// TIA Portal V21 export
// export: Created 2026-10-14T03:11:19.0543245Z, ExportSetting WithDefaults, DisplayName Totally Integrated Automation Portal, DisplayVersion V21, DisplayName STEP 7 Professional, DisplayVersion V21, DisplayName STEP 7 Safety, DisplayVersion V21, DisplayName Tech WebApplication, DisplayVersion V21, DisplayName WinCC Basic/Comfort/Advanced, DisplayVersion V21, DisplayName WinCC Unified, DisplayVersion V21
TagTable "PID_LCCA"
  LLCCA_PID_DB_Input : Real  (HMI_Connection_1, 100 ms)
  LLCCA_PID_DB_Out : Real  (HMI_Connection_1, 100 ms)
  LLCCA_PID_DB_Setpoint : Real  (HMI_Connection_1, 100 ms)
  LLCCA_PID_DB_ioKp : Real  (HMI_Connection_1, 1 s)
  LLCCA_PID_DB_ioTi : Real  (HMI_Connection_1, 1 s)
  LLCCA_PID_DB_ioTd : Real  (HMI_Connection_1, 1 s)
  LLCCA_PID_DB_Terms_p : Real  (HMI_Connection_1, 100 ms)
  LLCCA_PID_DB_Terms_i : Real  (HMI_Connection_1, 100 ms)
  LLCCA_PID_DB_Terms_d : Real  (HMI_Connection_1, 100 ms)
  LLCCA_PID_DB_statIntegralSum : Real  (HMI_Connection_1, 100 ms)
  LLCCA_PID_DB_statAdvanced_outMin : Real  (HMI_Connection_1, 1 s)
  LLCCA_PID_DB_statAdvanced_outMax : Real  (HMI_Connection_1, 1 s)
  LLCCA_PID_DB_statAdvanced_derivateFilter : Real  (HMI_Connection_1, 1 s)
  LLCCA_PID_DB_ioMode : USInt  (HMI_Connection_1, 100 ms)
  LLCCA_PID_DB_ManualValue : Real  (HMI_Connection_1, 1 s)
  LLCCA_PID_DB_statStepTuning_state : USInt  (HMI_Connection_1, 100 ms)
  LLCCA_PID_DB_statStepTuning_t : Real  (HMI_Connection_1, 100 ms)
  LLCCA_PID_DB_statAdvanced_inputFilter : Real  (HMI_Connection_1, 1 s)
  LLCCA_PID_DB_statAdvanced_tuningRule : USInt  (HMI_Connection_1, 1 s)
